Staubli VAL3: Data.dtx


